TYPE ST_Axis :
STRUCT
	stNcTOPLC: ST_NcTOPLC_AxisRef;
	stPLCTONC: ST_PLCTONC_AxisRef;
	stAxisStatus: ST_AxisStatus;
	stAxisParam: ST_AxisParameter;
	stCodToNCParam: ST_CodToNCParam;
END_STRUCT
END_TYPE

(* stored: Version 1.1.0.1, ProductVersion 3.1.4024.12
   DUT ST_Axis: Id {9c240aec-822f-47e2-81aa-9ec48fbc2df6} *)
